// TIA Portal V21 export
// export: Created 2026-11-11T00:47:31.314673Z, ExportSetting WithDefaults, DisplayName Totally Integrated Automation Portal, DisplayVersion V21 Update 3, DisplayName STEP 7 Professional, DisplayVersion V21 Update 3, DisplayName STEP 7 Safety, DisplayVersion V21, DisplayName Tech WebApplication, DisplayVersion V21, DisplayName WinCC Basic/Comfort/Advanced, DisplayVersion V21 Update 3, DisplayName WinCC Unified, DisplayVersion V21 Update 3
FUNCTION_BLOCK "FB_Fbd_ex120"   // FB131, FBD
{ S7_Optimized_Access := 'TRUE' }
VERSION : 0.1
// stored: AutoNumber true, IsIECCheckEnabled false, IsRetainMemResEnabled false, MemoryReserve 100, SetENOAutomatically false, UDAEnableTagReadback false
   VAR_INPUT
      v_alarm : ALARM_BASE;
   END_VAR
   VAR_OUTPUT
      v_alarmstate : Byte;
      v_error : Bool;
      v_status : Word;
   END_VAR
BEGIN

REGION Network 1: Get_AlarmState - Output alarm status
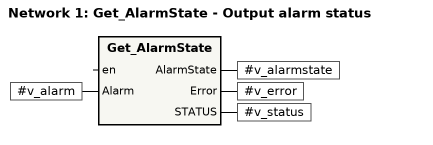
   Get_AlarmState(Alarm := #v_alarm, AlarmState => #v_alarmstate, Error => #v_error, STATUS => #v_status);
END_REGION
END_FUNCTION_BLOCK
